INTERFACE ITF_Blikjesband

METHOD Aborted : BOOL
VAR_INPUT
END_VAR
END_METHOD

METHOD Aborting : BOOL
VAR_INPUT
END_VAR
END_METHOD

METHOD Clearing : BOOL
VAR_INPUT
END_VAR
END_METHOD

METHOD Execute : BOOL
VAR_INPUT
END_VAR
END_METHOD

METHOD Held : BOOL
VAR_INPUT
END_VAR
END_METHOD

METHOD Holding : BOOL
VAR_INPUT
END_VAR
END_METHOD

METHOD Idle : BOOL
VAR_INPUT
END_VAR
END_METHOD

METHOD Resetting : BOOL
VAR_INPUT
END_VAR
END_METHOD

METHOD Starting : BOOL
VAR_INPUT
END_VAR
END_METHOD

METHOD Stopped : BOOL
VAR_INPUT
END_VAR
END_METHOD

METHOD Stopping : BOOL
VAR_INPUT
END_VAR
END_METHOD

METHOD Suspended : BOOL
VAR_INPUT
END_VAR
END_METHOD

METHOD Suspending : BOOL
VAR_INPUT
END_VAR
END_METHOD

METHOD Unholding : BOOL
VAR_INPUT
END_VAR
END_METHOD

METHOD Unsuspending : BOOL
VAR_INPUT
END_VAR
END_METHOD

END_INTERFACE

(* stored: Version 1.1.0.1
   Itf ITF_Blikjesband: Id {199bd5b4-7d2e-4c6e-ad31-02e50f35f66c}
   Folder Methods: Id {e8072a77-bb84-4c42-a35c-24150fa7685a}
   Method Aborted: Id {6620fa05-d309-424d-8d34-56a2b22d147c}
   Method Aborting: Id {ceedd066-ac35-478c-9e8f-b226e219f6d7}
   Method Clearing: Id {e636d0dc-c22e-4aba-a7e8-295d25822208}
   Method Execute: Id {ab09940a-6e45-4ff8-b1a4-9f3273b5b5cb}
   Method Held: Id {691941b4-400f-4b76-887f-ce7d6290d7e1}
   Method Holding: Id {6b32d497-022c-4820-9464-4d3ddecb7295}
   Method Idle: Id {a5541aeb-7b6c-46ec-a2da-2dc7edd094d5}
   Method Resetting: Id {da584811-c058-4791-a9eb-faaa1f98a9f7}
   Method Starting: Id {4c2a63eb-b3ac-4023-821b-177434e38342}
   Method Stopped: Id {7fc41be8-4ec9-42f2-9cf4-4754146f2185}
   Method Stopping: Id {3442d4d8-fdd5-4f4c-bd97-8aa97c68e92a}
   Method Suspended: Id {2869b93a-e4b5-4bf8-8777-2808abd2107d}
   Method Suspending: Id {f258df60-da31-4ae9-bb35-6555f570a650}
   Method Unholding: Id {42ec270f-b690-4808-8f74-025546006f3d}
   Method Unsuspending: Id {6c60b7e9-e51f-4fe5-b572-3ed555bb1762} *)
